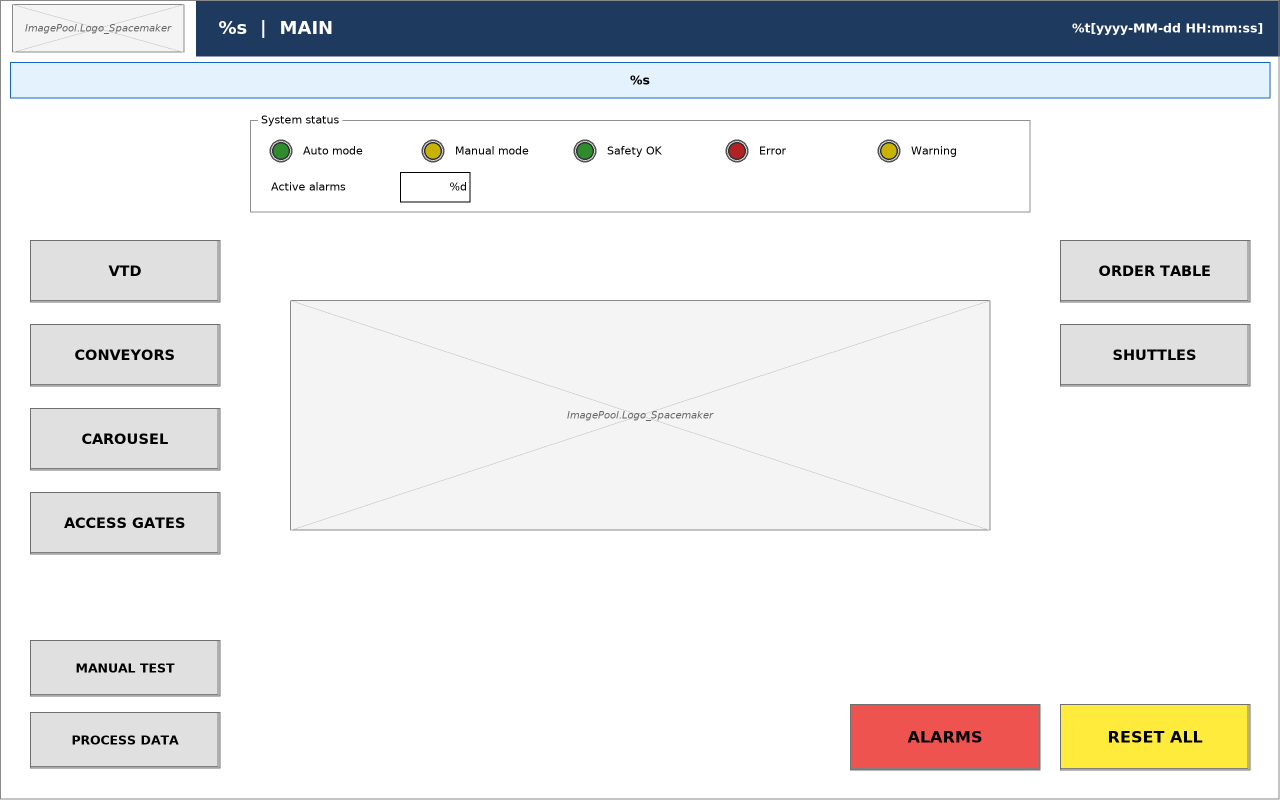
VISUALIZATION Main  // 1280x800
    Rectangle (0,0 196x56)
        OnMouseClick: change screen: Main
    Image (12,4 172x48), image: ImagePool.Logo_Spacemaker
        OnMouseClick: change screen: Main
    Rectangle (196,0 1084x56), "%s | MAIN", text variable: GVL_HMI_System.stStatus.sSystemName
    Rectangle (930,8 336x40), "%t[yyyy-MM-dd HH:mm:ss]", text variable: GVL_HMI_System.stStatus.dtNow
    Rectangle (10,62 1260x36), "%s", text variable: GVL_HMI_System.stStatus.sMessage, colour toggle: GVL_HMI_System.stStatus.bMessageAlarm
    GroupBox (250,112 780x100), "System status"
    Lamp1 (268,138 26x26), variable: GVL_HMI_System.stStatus.bAutoMode, style: Lamp-Lamp1-Green
    Rectangle (300,136 112x30), "Auto mode"
    Lamp1 (420,138 26x26), variable: GVL_HMI_System.stStatus.bManualMode, style: Lamp-Lamp1-Yellow
    Rectangle (452,136 112x30), "Manual mode"
    Lamp1 (572,138 26x26), variable: GVL_HMI_System.stStatus.bSafetyOk, style: Lamp-Lamp1-Green
    Rectangle (604,136 112x30), "Safety OK"
    Lamp1 (724,138 26x26), variable: GVL_HMI_System.stStatus.bError, style: Lamp-Lamp1-Red
    Rectangle (756,136 112x30), "Error"
    Lamp1 (876,138 26x26), variable: GVL_HMI_System.stStatus.bWarning, style: Lamp-Lamp1-Yellow
    Rectangle (908,136 112x30), "Warning"
    Rectangle (268,172 130x30), "Active alarms"
    Rectangle (400,172 70x30), "%d", text variable: GVL_HMI_System.stStatus.uiActiveAlarms
    Image (290,300 700x230), image: ImagePool.Logo_Spacemaker
    Button (30,240 190x62), "VTD", colour toggle: GVL_HMI_System.stVtd.stSummary.bError
        OnMouseClick: change screen: VTD
    Button (30,324 190x62), "CONVEYORS"
        OnMouseClick: change screen: CNV
    Button (30,408 190x62), "CAROUSEL"
        OnMouseClick: change screen: Carrousel
    Button (30,492 190x62), "ACCESS GATES"
        OnMouseClick: change screen: Access_Gates
    Button (30,640 190x56), "MANUAL TEST"
        OnMouseClick: change screen: VTDManualTest
    Button (30,712 190x56), "PROCESS DATA"
        OnMouseClick: change screen: Visualization
    Button (1060,240 190x62), "ORDER TABLE"
        OnMouseClick: change screen: Order_Table
    Button (1060,324 190x62), "SHUTTLES"
        OnMouseClick: change screen: Shuttles
    Button (850,704 190x66), "ALARMS"
        OnMouseClick: change screen: Alarms
    Button (1060,704 190x66), "RESET ALL"
        tap GVL_HMI_System.stCommand.bResetAll p3779583253=TRUE
END_VISUALIZATION

(* stored: Version 1.1.0.1
   Visu Main: Id {3055a09b-9538-4080-8201-d34ec6b675c3} *)
